(* IEC 61131-3 sources: plc-process-lib/tests/POUs/Helpers/FB_FopdtModel, 3 files *)

(* ---- FB_FopdtModel.decl.st ---- *)
// Назначение: модель объекта «первый порядок + запаздывание» (FOPDT) для тестов ПИД в замкнутом
//             контуре: y[k+1] = y[k] + dt/T·(K·u[k - L/dt] - y[k]), шаг dt = 0,1 с, запаздывание
//             L = 4 с — кольцо на 40 отсчётов (контракт API.md, 22.5 и 23.1). Состояние — LREAL,
//             выход rY — REAL. Шаг модели — метод Step; тело пустое. Эталон —
//             tools/reference/pid.py, класс Fopdt. Параметры объекта вымышленные. Только для тестов.
// Автор:      kr0nsch
// Версия:     0.1.0
// Документ:   docs/fb/FB_PID.md, раздел «Тесты»
FUNCTION_BLOCK FB_FopdtModel
VAR CONSTANT
    DT_S        : LREAL := 0.1;   // шаг модели, с
    RING_SIZE   : UINT := 40;     // длина кольца = запаздывание в шагах: L / dt = 4 с / 0,1 с
END_VAR
VAR_INPUT
    rU_pct : REAL;                // вход объекта (выход регулятора), %
    rGain  : REAL := 2.0;         // K, инж. ед. на %
    rT_s   : REAL := 20.0;        // T, с
END_VAR
VAR_OUTPUT
    rY : REAL;                    // выход объекта, инж. ед.
END_VAR
VAR
    arDelay : ARRAY[0..RING_SIZE - 1] OF REAL;   // кольцо запаздывания
    uiHead  : UINT;                   // самая старая запись кольца: u[k - 40]
    lrY     : LREAL;                  // состояние y
END_VAR

(* ---- Step.method.decl.st ---- *)
// Один шаг модели dt = 0,1 с: из кольца берётся вход 40 шагов назад, на его место пишется rU_pct
METHOD PUBLIC Step
VAR
    rUDelayed : REAL;   // u[k - 40]
END_VAR

(* ---- Step.method.impl.st ---- *)
rUDelayed := arDelay[uiHead];
arDelay[uiHead] := rU_pct;
uiHead := uiHead + 1;
IF uiHead >= RING_SIZE THEN
    uiHead := 0;
END_IF
lrY := lrY + DT_S / REAL_TO_LREAL(rT_s) * (REAL_TO_LREAL(rGain) * REAL_TO_LREAL(rUDelayed) - lrY);
rY := LREAL_TO_REAL(lrY);
